// Core S3.12 - the SET result, valid on Done.
TYPE ST_AnalogOutputOutCmd :
STRUCT
    Applied : LREAL;
END_STRUCT
END_TYPE

(* stored: Version 1.1.0.1, ProductVersion 3.1.4024.12
   DUT ST_AnalogOutputOutCmd: Id {8c7983f6-7d8c-4ba9-9687-b37c76077132} *)
